% RSLogix 500 project PROGRAM 5.RSS, saved by version 8.30.00.16 %
PROJECT "UNTITLED"    % processor: Bul.1763 MicroLogix 1100 Series B %

PROGRAM FILES
  LAD 2 "MAIN"  2 rungs
  LAD 4 "PROC_LOGIC"  6 rungs

DATA FILES
  O0 OUTPUT  4 elements
  I1 INPUT  6 elements
  S2 STATUS  66 elements
  B3 BINARY  1 elements
  T4 TIMER  2 elements
  C5 COUNTER  1 elements
  R6 CONTROL  1 elements
  N7 INTEGER  1 elements
  F8 FLOAT  3 elements

LADDER 2 "MAIN"
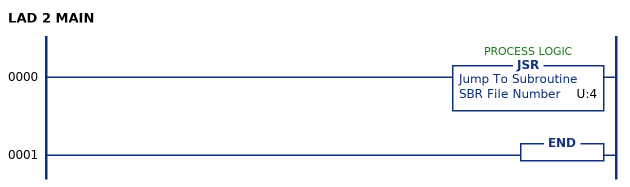
% Rung: 0 %
SOR JSR U:4 EOR
%   U:4  "PROCESS LOGIC" %
% Rung: 1 %
SOR END EOR

LADDER 4 "PROC_LOGIC"
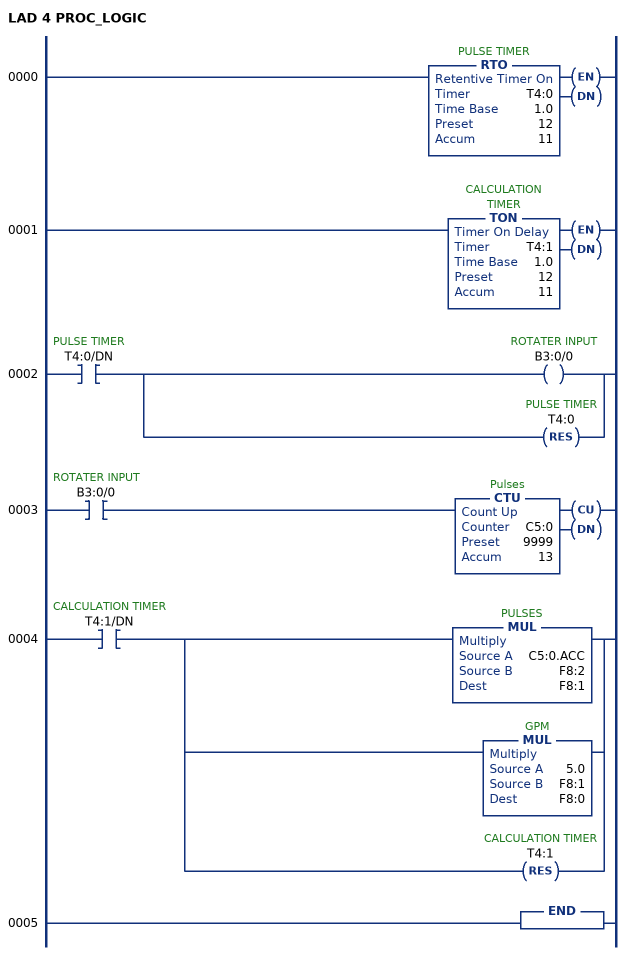
% Rung: 0 %
SOR RTO T4:0 1.0 12 11 EOR
%   T4:0  "PULSE TIMER" %
% Rung: 1 %
SOR TON T4:1 1.0 12 11 EOR
%   T4:1  "CALCULATION TIMER" %
% Rung: 2 %
SOR XIC T4:0/DN BST OTE B3:0/0 NXB RES T4:0 BND EOR
%   T4:0  "PULSE TIMER" %
%   B3:0/0  "ROTATER INPUT" %
% Rung: 3 %
SOR XIC B3:0/0 CTU C5:0 9999 13 EOR
%   B3:0/0  "ROTATER INPUT" %
%   C5:0  "Pulses" %
% Rung: 4 %
SOR XIC T4:1/DN BST MUL C5:0.ACC F8:2 F8:1 NXB MUL 5.0 F8:1 F8:0 NXB RES T4:1 BND EOR
%   T4:1  "CALCULATION TIMER" %
%   C5:0.ACC  "PULSES ACCUMUILATIONS" %
%   F8:2  "k-factor" %
%   F8:1  PULSES %
%   F8:0  "GPM" %
% Rung: 5 %
SOR END EOR

OTHER DOCUMENTED ADDRESSES
  B3:0/1  "ONS"
  U:3  "IO"

DATA TABLE (non-zero values as saved)
DATA T4
% .PRE .ACC %
% T4:0 % 12 11
% T4:1 % 12 11
DATA C5
% .PRE .ACC %
% C5:0 % 9999 13
DATA F8
% F8:0 % 409.5 81.9 6.3
